// LS Electric XG5000 project: NewProject
// PLC LSPLC

PROGRAM NewProgram (task: 스캔 프로그램)

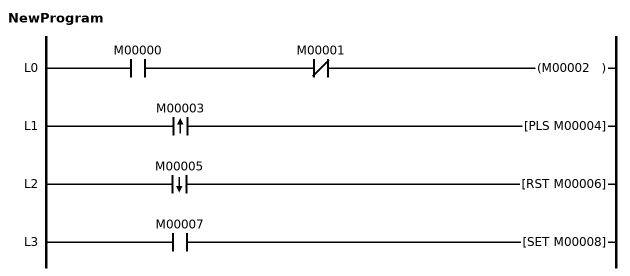
; L0
LOAD      M00000
AND NOT   M00001
OUT       M00002
; L1
LOADP     M00003
OUTP      M00004
; L2
LOADN     M00005
RST       M00006
; L3
LOAD      M00007
SET       M00008